(* PLC project TBEN_L5_PLC11.project, CODESYS CODESYS V3.5 SP21 Patch 1 *)
(* stored: creationDateTime 2026-11-07T15:35:09.2062848, modificationDateTime 2026-11-07T15:09:07.4034196 *)

// Trừu tượng hoá đọc/ghi record PROFINET (CommFB.WRREC/RDREC thật hoặc mock Simulation)
// Quy ước như CommFB: giữ xReq = TRUE tới khi có kết quả, hạ xReq ít nhất 1 lần gọi trước request mới; gọi mỗi chu kỳ đúng 1 lần.
INTERFACE ITF_IolRecordAccess
// Ghi record (WRREC). Trả TRUE khi đã kết thúc (xDone hoặc xError).
METHOD Write : BOOL
VAR_INPUT
    xReq   : BOOL;
    dwId   : DWORD;                 // ID submodule (CommFB.SUBSLOT_ID), mock bỏ qua
    iIndex : INT;                   // record index (0xB400 truyền dạng INT)
    iLen   : INT;                   // số byte ghi
    pData  : POINTER TO BYTE;
END_VAR
VAR_OUTPUT
    xDone    : BOOL;
    xBusy    : BOOL;
    xError   : BOOL;
    dwStatus : DWORD;               // STATUS PNIO 4 byte
END_VAR
END_METHOD
// Đọc record (RDREC). Trả TRUE khi đã kết thúc (xValid hoặc xError).
METHOD Read : BOOL
VAR_INPUT
    xReq   : BOOL;
    dwId   : DWORD;
    iIndex : INT;
    iMLen  : INT;                   // kích thước buffer nhận
    pData  : POINTER TO BYTE;
END_VAR
VAR_OUTPUT
    xValid   : BOOL;
    xBusy    : BOOL;
    xError   : BOOL;
    dwStatus : DWORD;
    iLen     : INT;                 // số byte nhận được
END_VAR
END_METHOD
END_INTERFACE
